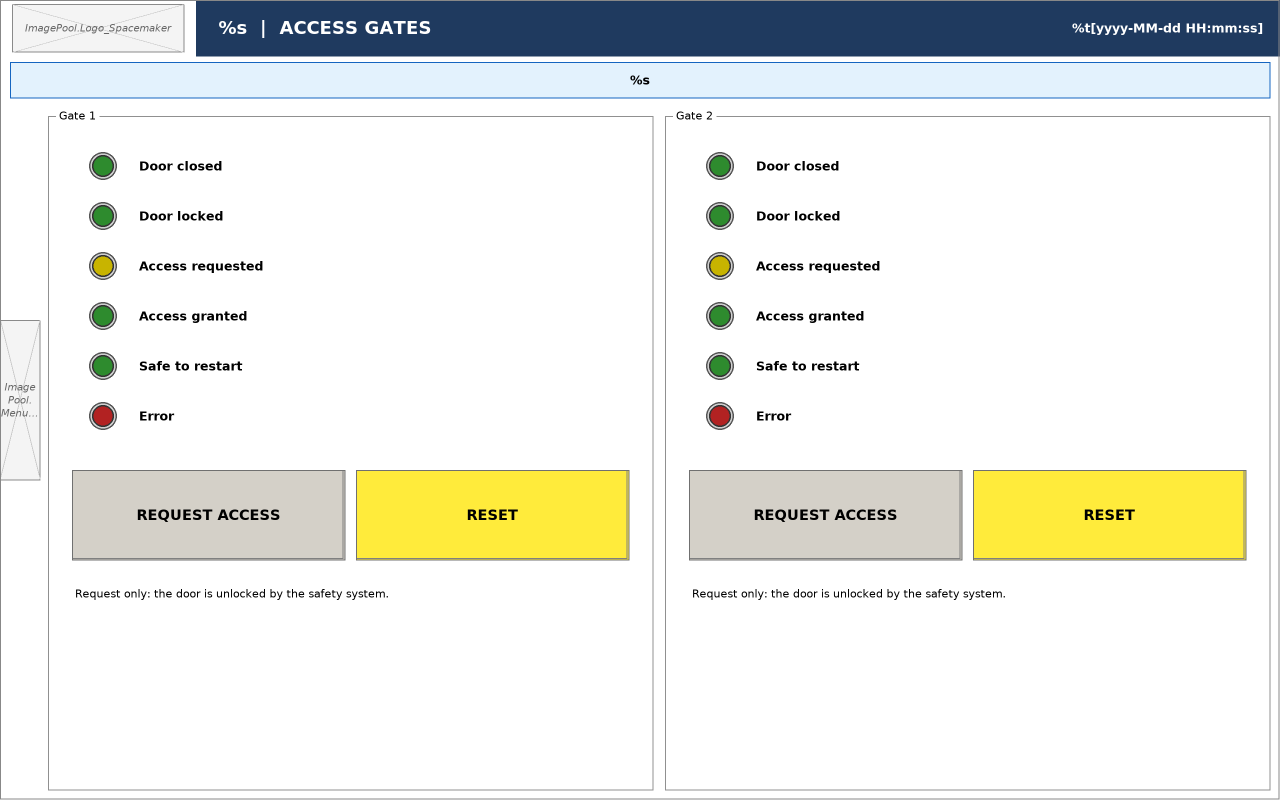
VISUALIZATION Access_Gates  // 1280x800
    Rectangle (0,0 196x56)
        OnMouseClick: change screen: Main
    Image (12,4 172x48), image: ImagePool.Logo_Spacemaker
        OnMouseClick: change screen: Main
    Rectangle (196,0 1084x56), "%s | ACCESS GATES", text variable: GVL_HMI_System.stStatus.sSystemName
    Rectangle (930,8 336x40), "%t[yyyy-MM-dd HH:mm:ss]", text variable: GVL_HMI_System.stStatus.dtNow
    Rectangle (10,62 1260x36), "%s", text variable: GVL_HMI_System.stStatus.sMessage, colour toggle: GVL_HMI_System.stStatus.bMessageAlarm
    GroupBox (48,108 605x682), "Gate 1"
    Lamp1 (87,150 32x32), variable: GVL_HMI_Gates.astGate[1].bClosed, style: Lamp-Lamp1-Green
    Rectangle (136,150 356x32), "Door closed"
    Lamp1 (87,200 32x32), variable: GVL_HMI_Gates.astGate[1].bLocked, style: Lamp-Lamp1-Green
    Rectangle (136,200 356x32), "Door locked"
    Lamp1 (87,250 32x32), variable: GVL_HMI_Gates.astGate[1].bAccessRequested, style: Lamp-Lamp1-Yellow
    Rectangle (136,250 356x32), "Access requested"
    Lamp1 (87,300 32x32), variable: GVL_HMI_Gates.astGate[1].bAccessGranted, style: Lamp-Lamp1-Green
    Rectangle (136,300 356x32), "Access granted"
    Lamp1 (87,350 32x32), variable: GVL_HMI_Gates.astGate[1].bSafeToRestart, style: Lamp-Lamp1-Green
    Rectangle (136,350 356x32), "Safe to restart"
    Lamp1 (87,400 32x32), variable: GVL_HMI_Gates.astGate[1].bError, style: Lamp-Lamp1-Red
    Rectangle (136,400 356x32), "Error"
    Button (72,470 273x90), "REQUEST ACCESS"
        tap GVL_HMI_Gates.astCommand[1].bRequestAccess p3779583253=TRUE
    Button (356,470 273x90), "RESET"
        tap GVL_HMI_Gates.astCommand[1].bReset p3779583253=TRUE
    Rectangle (72,580 557x28), "Request only: the door is unlocked by the safety system."
    GroupBox (665,108 605x682), "Gate 2"
    Lamp1 (704,150 32x32), variable: GVL_HMI_Gates.astGate[2].bClosed, style: Lamp-Lamp1-Green
    Rectangle (753,150 356x32), "Door closed"
    Lamp1 (704,200 32x32), variable: GVL_HMI_Gates.astGate[2].bLocked, style: Lamp-Lamp1-Green
    Rectangle (753,200 356x32), "Door locked"
    Lamp1 (704,250 32x32), variable: GVL_HMI_Gates.astGate[2].bAccessRequested, style: Lamp-Lamp1-Yellow
    Rectangle (753,250 356x32), "Access requested"
    Lamp1 (704,300 32x32), variable: GVL_HMI_Gates.astGate[2].bAccessGranted, style: Lamp-Lamp1-Green
    Rectangle (753,300 356x32), "Access granted"
    Lamp1 (704,350 32x32), variable: GVL_HMI_Gates.astGate[2].bSafeToRestart, style: Lamp-Lamp1-Green
    Rectangle (753,350 356x32), "Safe to restart"
    Lamp1 (704,400 32x32), variable: GVL_HMI_Gates.astGate[2].bError, style: Lamp-Lamp1-Red
    Rectangle (753,400 356x32), "Error"
    Button (689,470 273x90), "REQUEST ACCESS"
        tap GVL_HMI_Gates.astCommand[2].bRequestAccess p3779583253=TRUE
    Button (973,470 273x90), "RESET"
        tap GVL_HMI_Gates.astCommand[2].bReset p3779583253=TRUE
    Rectangle (689,580 557x28), "Request only: the door is unlocked by the safety system."
    Rectangle (0,320 40x160)
        OnMouseEnter: OpenDialog Dialog=Dialog, OpenModal=True, PositionX=0, PositionY=0
        OnMouseClick: OpenDialog Dialog=Dialog, OpenModal=True, PositionX=0, PositionY=0
    Image (0,320 40x160), image: ImagePool.Menu_Tab
        OnMouseEnter: OpenDialog Dialog=Dialog, OpenModal=True, PositionX=0, PositionY=0
        OnMouseClick: OpenDialog Dialog=Dialog, OpenModal=True, PositionX=0, PositionY=0
END_VISUALIZATION

(* stored: Version 1.1.0.1
   Visu Access_Gates: Id {01892bde-30c2-44b5-aa78-ae2fd3431384} *)
